FUNCTION_BLOCK FB_SimAxis
VAR_OUTPUT
    PositionMm : DINT;
END_VAR

METHOD MoveToward : BOOL
VAR_INPUT
    TargetMm : DINT;
    MaxStepMm : DINT;
END_VAR
// Deterministic virtual axis. One invocation corresponds to one 10 ms task tick.
PositionMm := PositionMm + LIMIT(-MaxStepMm, TargetMm - PositionMm, MaxStepMm);
MoveToward := PositionMm = TargetMm;
END_METHOD

METHOD Home
PositionMm := 0;
END_METHOD

END_FUNCTION_BLOCK

(* stored: Version 1.1.0.1
   POU FB_SimAxis: Id {69468DC3-8A7A-45D7-9465-000000000001}
   Method MoveToward: Id {69468DC3-8A7A-45D7-9465-000000000002}
   Method Home: Id {69468DC3-8A7A-45D7-9465-000000000003} *)
